SUBAPPLICATION Heckschieber (* Subapplication Type *)
  (* Standard: 61499-2 *)
  (* Version 1.0, 2023-01-29, Franz *)
  IMPORT DefaultPool::SoftKey_Heckschieber;
  IMPORT isobus::UT::io::Softkey::SoftKeyActivationCode::SK_RELEASED;
  IMPORT DefaultPool::AuxInput_Heckschieber;
  IMPORT isobus::UT::io::Auxiliary::IN::AuxiliaryState::AuxDisabled;
  IMPORT DataPanel::io::MI::DQ::DataPanel_MI_DO::DigitalOutput_6B;
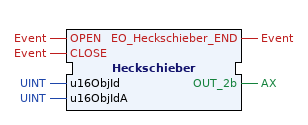
  EVENT_INPUT
    OPEN;
    CLOSE;
  END_EVENT
  EVENT_OUTPUT
    EO_Heckschieber_END;
  END_EVENT
  VAR_INPUT
    u16ObjId : UINT;
    u16ObjIdA : UINT;
  END_VAR
  PLUGS
    OUT_2b : adapter::types::unidirectional::AX;
  END_PLUGS
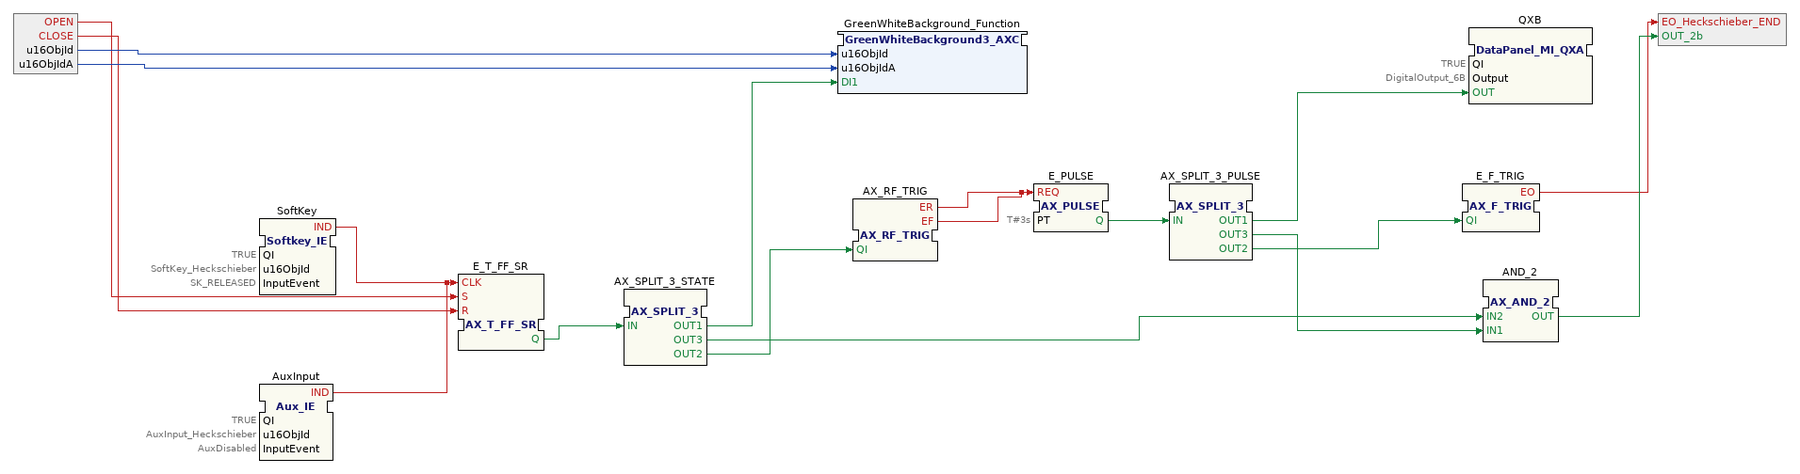
  FBS
    E_F_TRIG : adapter::events::unidirectional::AX_F_TRIG;
    QXB : DataPanel::io::MI::DQ::DataPanel_MI_QXA(QI := TRUE, Output := DigitalOutput_6B);
    E_T_FF_SR : adapter::events::unidirectional::AX_T_FF_SR;
    AX_SPLIT_3_STATE : adapter::events::unidirectional::AX_SPLIT_3;
    AX_RF_TRIG : adapter::events::unidirectional::AX_RF_TRIG;
    AX_SPLIT_3_PULSE : adapter::events::unidirectional::AX_SPLIT_3;
    AND_2 : adapter::booleanOperators::AX_AND_2;
    E_PULSE : adapter::events::unidirectional::timers::AX_PULSE(PT := T#3s);
    SoftKey : isobus::UT::io::Softkey::Softkey_IE(QI := TRUE, u16ObjId := SoftKey_Heckschieber, InputEvent := SK_RELEASED);
    AuxInput : isobus::UT::io::Auxiliary::IN::Aux_IE(QI := TRUE, u16ObjId := AuxInput_Heckschieber, InputEvent := AuxDisabled);
  END_FBS
  SUBAPPS
    GreenWhiteBackground_Function : MyLib::sys::GreenWhiteBackground3_AXC;
  END_SUBAPPS
  EVENT_CONNECTIONS
    E_F_TRIG.EO TO EO_Heckschieber_END;
    SoftKey.IND TO E_T_FF_SR.CLK;
    AuxInput.IND TO E_T_FF_SR.CLK;
    OPEN TO E_T_FF_SR.S;
    CLOSE TO E_T_FF_SR.R;
    AX_RF_TRIG.ER TO E_PULSE.REQ;
    AX_RF_TRIG.EF TO E_PULSE.REQ;
  END_CONNECTIONS
  DATA_CONNECTIONS
    u16ObjId TO GreenWhiteBackground_Function.u16ObjId;
    u16ObjIdA TO GreenWhiteBackground_Function.u16ObjIdA;
  END_CONNECTIONS
  ADAPTER_CONNECTIONS
    E_T_FF_SR.Q TO AX_SPLIT_3_STATE.IN;
    AX_SPLIT_3_STATE.OUT1 TO GreenWhiteBackground_Function.DI1;
    AX_SPLIT_3_STATE.OUT3 TO AND_2.IN2;
    E_PULSE.Q TO AX_SPLIT_3_PULSE.IN;
    AX_SPLIT_3_PULSE.OUT1 TO QXB.OUT;
    AX_SPLIT_3_PULSE.OUT3 TO AND_2.IN1;
    AND_2.OUT TO OUT_2b;
    AX_SPLIT_3_STATE.OUT2 TO AX_RF_TRIG.QI;
    AX_SPLIT_3_PULSE.OUT2 TO E_F_TRIG.QI;
  END_CONNECTIONS
END_SUBAPPLICATION
